(* IEC 61131-3 sources: kns-port-domestic/tools/port_metrics_tests/fixtures/app/src/POUs/FB_Pump, 3 files *)

(* ---- FB_Pump.decl.st ---- *)
// Насос: пример для метрик переноса
FUNCTION_BLOCK FB_Pump EXTENDS FB_Base
VAR_INPUT
    xStart : BOOL;
    stCfg : ST_PumpCfg;
END_VAR
VAR_OUTPUT
    xRunning : BOOL;
END_VAR
VAR
    tonDelay : TON;
END_VAR

(* ---- FB_Pump.impl.st ---- *)
SUPER^();
tonDelay(IN := xStart, PT := stCfg.tStartDelay);
xRunning := tonDelay.Q AND NOT xFault;
IF xRunning THEN
    Start();
ELSE
    Stop();
END_IF

(* ---- Start.method.decl.st ---- *)
METHOD Start : BOOL
VAR_INPUT
END_VAR
